Fanuc KAREL source: KC00036.KL

PROGRAM KC00036
%NOLOCKGROUP
%ENVIRONMENT KCLOP
VAR
  I: INTEGER
  J: INTEGER
  K: INTEGER
  R: REAL
  B: BOOLEAN
  S: STRING[80]
  T: STRING[80]
  P: PATH
  Q: PATH
  AI: ARRAY[8] OF INTEGER
  AB: ARRAY[244] OF BYTE
BEGIN
  I = KCL_STATUS
END KC00036
